TYPE ST_EL4022 :
STRUCT
    sTerminalName : STRING(80) := 'EL4022 | 2-Channel Analog Output 4..20mA';
    iEL4028_Ch1 AT %Q* : INT;
    iEL4028_Ch2 AT %Q* : INT;
    stTerminalInfo : ST_Terminal_Info;
END_STRUCT
END_TYPE

(* stored: Version 1.1.0.1, ProductVersion 3.1.4026.18
   DUT ST_EL4022: Id {b1541fe2-44f3-47f6-a421-e35168597bf4} *)
